(* Logix 5000 project; controller CIP vendor 1 type 14 code 106 rev 20.12; software revision 20.06; part 5 of 13 *)
(* tags used below, declared in another part *)
   Alarm_Ack : INT[8];
   Alarm_Present : INT[8];
   Alarm_Timer : TIMER[128];
   Bit : BOOL[128];
   IN_N7_100_199 : INT[100];
   Integer : DINT[150];
   OpCode_Pin : DINT[5];
   Recipe : RECIPE[41];
   RotaryONS : DINT;
   SCLD_Supply_Flow : REAL;
   SCLD_Supply_Pressure : REAL;
   SCLD_Wash_Chamber_Lvl : REAL;
   WashChamberDoorGasketCTRL : DINT;
(* MainProgram, continued *)

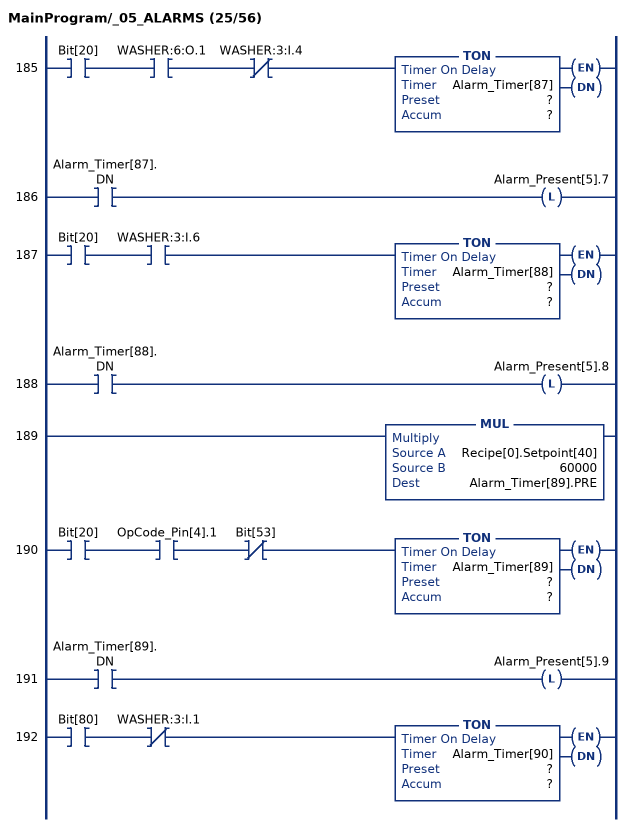
   [picture p67: MainProgram/_05_ALARMS rungs 185-192]
   185: XIC(Bit[20])XIC(WASHER:6:O.1)XIO(WASHER:3:I.4)TON(Alarm_Timer[87],?,?);
   186: XIC(Alarm_Timer[87].DN)OTL(Alarm_Present[5].7);
   187: XIC(Bit[20])XIC(WASHER:3:I.6)TON(Alarm_Timer[88],?,?);
   188: XIC(Alarm_Timer[88].DN)OTL(Alarm_Present[5].8);
   189: MUL(Recipe[0].Setpoint[40],60000,Alarm_Timer[89].PRE);
   190: XIC(Bit[20])XIC(OpCode_Pin[4].1)XIO(Bit[53])TON(Alarm_Timer[89],?,?);
   191: XIC(Alarm_Timer[89].DN)OTL(Alarm_Present[5].9);
   192: XIC(Bit[80])XIO(WASHER:3:I.1)TON(Alarm_Timer[90],?,?);
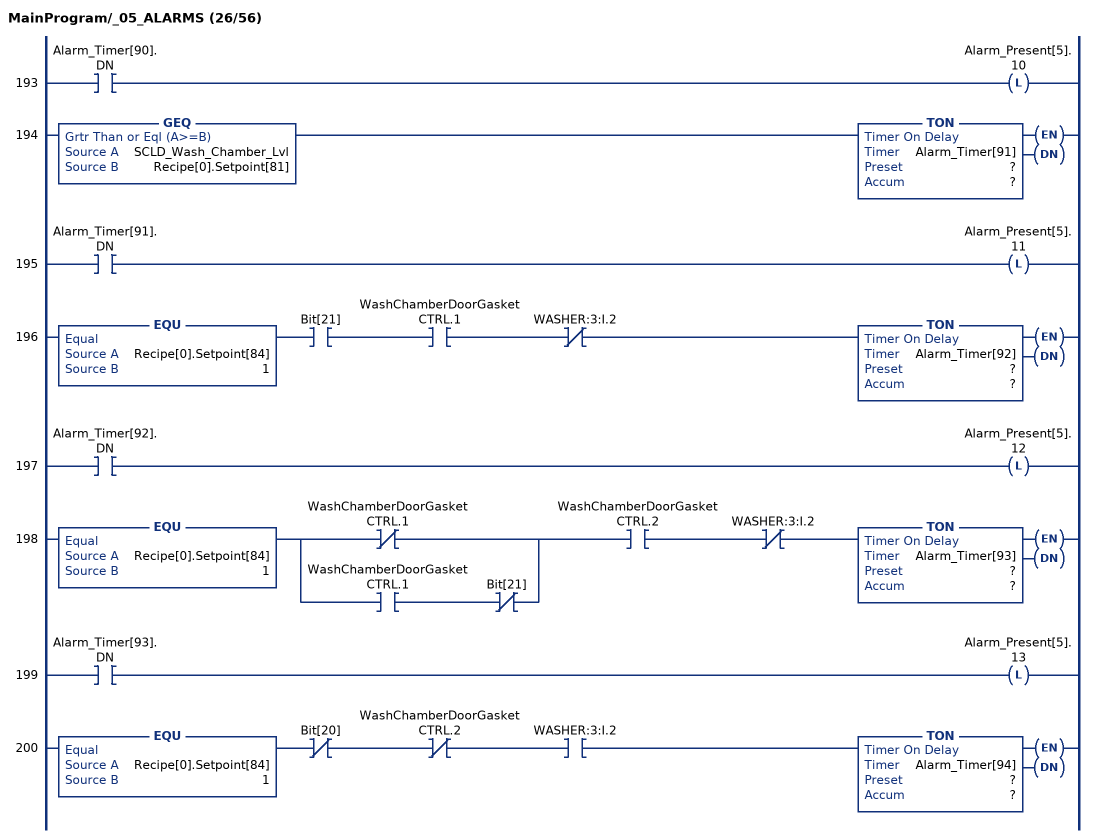
   193: XIC(Alarm_Timer[90].DN)OTL(Alarm_Present[5].10);
   194: GEQ(SCLD_Wash_Chamber_Lvl,Recipe[0].Setpoint[81])TON(Alarm_Timer[91],?,?);
   195: XIC(Alarm_Timer[91].DN)OTL(Alarm_Present[5].11);
   196: EQU(Recipe[0].Setpoint[84],1)XIC(Bit[21])XIC(WashChamberDoorGasketCTRL.1)XIO(WASHER:3:I.2)TON(Alarm_Timer[92],?,?);
   197: XIC(Alarm_Timer[92].DN)OTL(Alarm_Present[5].12);
   198: EQU(Recipe[0].Setpoint[84],1)[XIO(WashChamberDoorGasketCTRL.1) ,XIC(WashChamberDoorGasketCTRL.1) XIO(Bit[21]) ]XIC(WashChamberDoorGasketCTRL.2)XIO(WASHER:3:I.2)TON(Alarm_Timer[93],?,?);
   199: XIC(Alarm_Timer[93].DN)OTL(Alarm_Present[5].13);
   200: EQU(Recipe[0].Setpoint[84],1)XIO(Bit[20])XIO(WashChamberDoorGasketCTRL.2)XIC(WASHER:3:I.2)TON(Alarm_Timer[94],?,?);
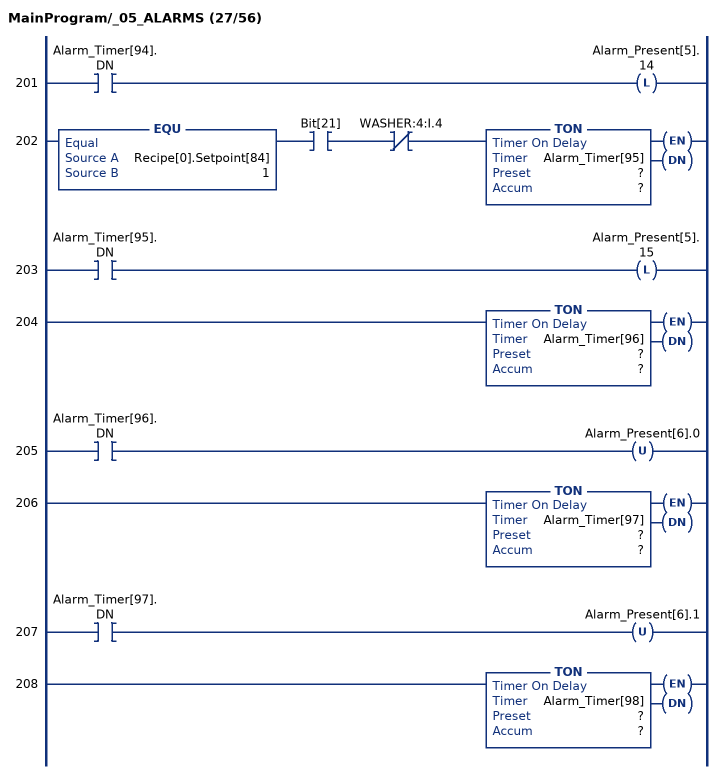
   201: XIC(Alarm_Timer[94].DN)OTL(Alarm_Present[5].14);
   202: EQU(Recipe[0].Setpoint[84],1)XIC(Bit[21])XIO(WASHER:4:I.4)TON(Alarm_Timer[95],?,?);
   203: XIC(Alarm_Timer[95].DN)OTL(Alarm_Present[5].15);
   204: TON(Alarm_Timer[96],?,?);
   205: XIC(Alarm_Timer[96].DN)OTU(Alarm_Present[6].0);
   206: TON(Alarm_Timer[97],?,?);
   207: XIC(Alarm_Timer[97].DN)OTU(Alarm_Present[6].1);
   208: TON(Alarm_Timer[98],?,?);
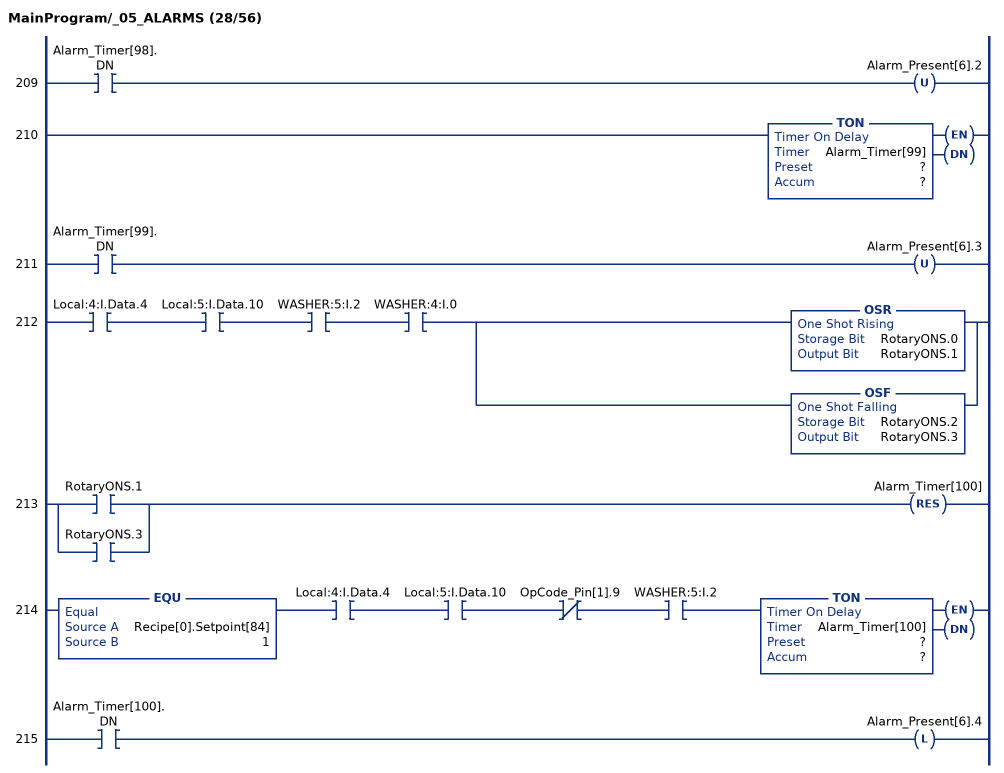
   209: XIC(Alarm_Timer[98].DN)OTU(Alarm_Present[6].2);
   210: TON(Alarm_Timer[99],?,?);
   211: XIC(Alarm_Timer[99].DN)OTU(Alarm_Present[6].3);
   212: XIC(Local:4:I.Data.4)XIC(Local:5:I.Data.10)XIC(WASHER:5:I.2)XIC(WASHER:4:I.0)[OSR(RotaryONS.0,RotaryONS.1) ,OSF(RotaryONS.2,RotaryONS.3) ];
   213: [XIC(RotaryONS.1) ,XIC(RotaryONS.3) ]RES(Alarm_Timer[100]);
   214: EQU(Recipe[0].Setpoint[84],1)XIC(Local:4:I.Data.4)XIC(Local:5:I.Data.10)XIO(OpCode_Pin[1].9)XIC(WASHER:5:I.2)TON(Alarm_Timer[100],?,?);
   215: XIC(Alarm_Timer[100].DN)OTL(Alarm_Present[6].4);
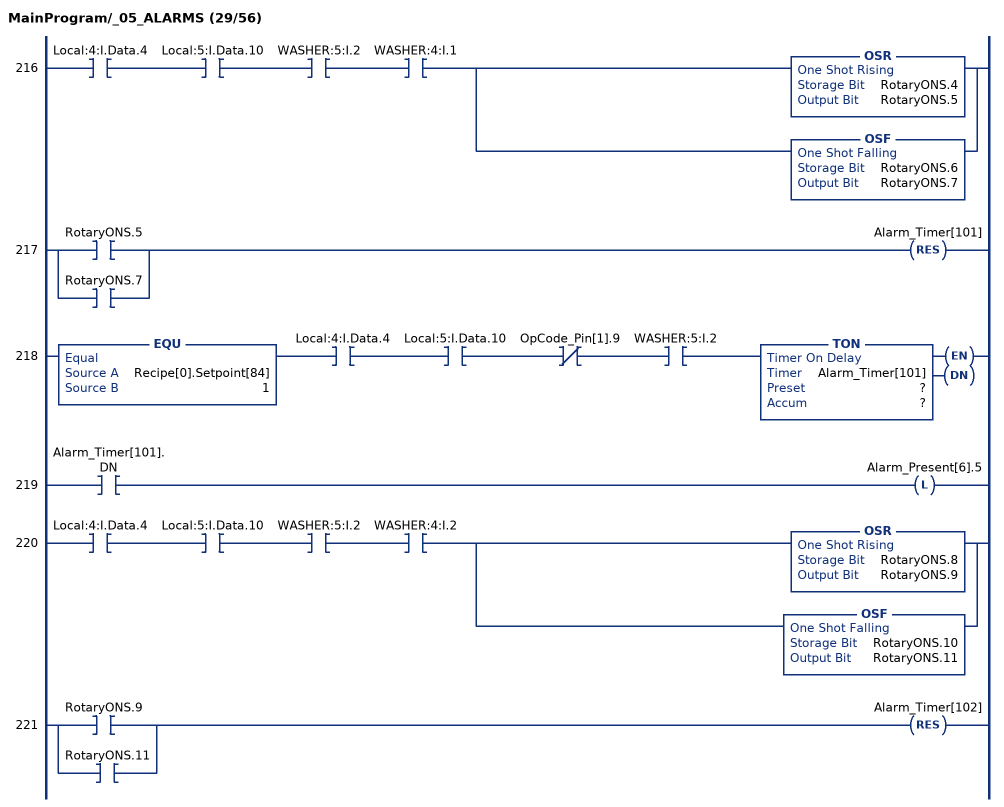
   216: XIC(Local:4:I.Data.4)XIC(Local:5:I.Data.10)XIC(WASHER:5:I.2)XIC(WASHER:4:I.1)[OSR(RotaryONS.4,RotaryONS.5) ,OSF(RotaryONS.6,RotaryONS.7) ];
   217: [XIC(RotaryONS.5) ,XIC(RotaryONS.7) ]RES(Alarm_Timer[101]);
   218: EQU(Recipe[0].Setpoint[84],1)XIC(Local:4:I.Data.4)XIC(Local:5:I.Data.10)XIO(OpCode_Pin[1].9)XIC(WASHER:5:I.2)TON(Alarm_Timer[101],?,?);
   219: XIC(Alarm_Timer[101].DN)OTL(Alarm_Present[6].5);
   220: XIC(Local:4:I.Data.4)XIC(Local:5:I.Data.10)XIC(WASHER:5:I.2)XIC(WASHER:4:I.2)[OSR(RotaryONS.8,RotaryONS.9) ,OSF(RotaryONS.10,RotaryONS.11) ];
   221: [XIC(RotaryONS.9) ,XIC(RotaryONS.11) ]RES(Alarm_Timer[102]);
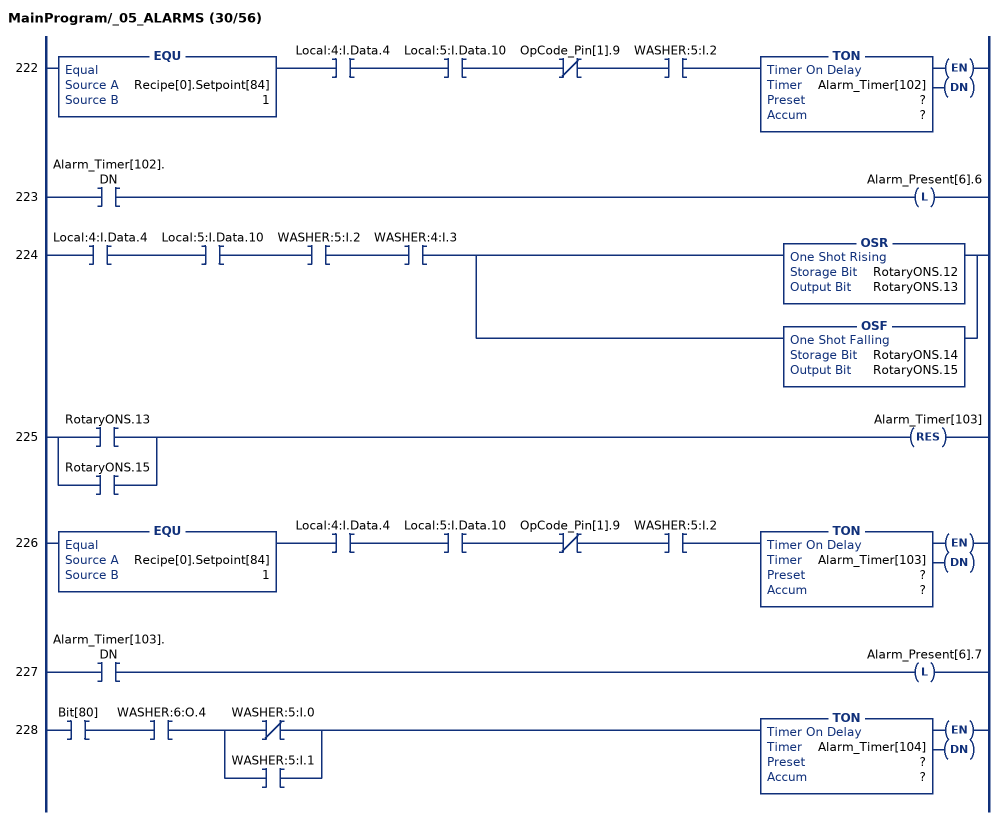
   222: EQU(Recipe[0].Setpoint[84],1)XIC(Local:4:I.Data.4)XIC(Local:5:I.Data.10)XIO(OpCode_Pin[1].9)XIC(WASHER:5:I.2)TON(Alarm_Timer[102],?,?);
   223: XIC(Alarm_Timer[102].DN)OTL(Alarm_Present[6].6);
   224: XIC(Local:4:I.Data.4)XIC(Local:5:I.Data.10)XIC(WASHER:5:I.2)XIC(WASHER:4:I.3)[OSR(RotaryONS.12,RotaryONS.13) ,OSF(RotaryONS.14,RotaryONS.15) ];
   225: [XIC(RotaryONS.13) ,XIC(RotaryONS.15) ]RES(Alarm_Timer[103]);
   226: EQU(Recipe[0].Setpoint[84],1)XIC(Local:4:I.Data.4)XIC(Local:5:I.Data.10)XIO(OpCode_Pin[1].9)XIC(WASHER:5:I.2)TON(Alarm_Timer[103],?,?);
   227: XIC(Alarm_Timer[103].DN)OTL(Alarm_Present[6].7);
   228: XIC(Bit[80])XIC(WASHER:6:O.4)[XIO(WASHER:5:I.0) ,XIC(WASHER:5:I.1) ]TON(Alarm_Timer[104],?,?);
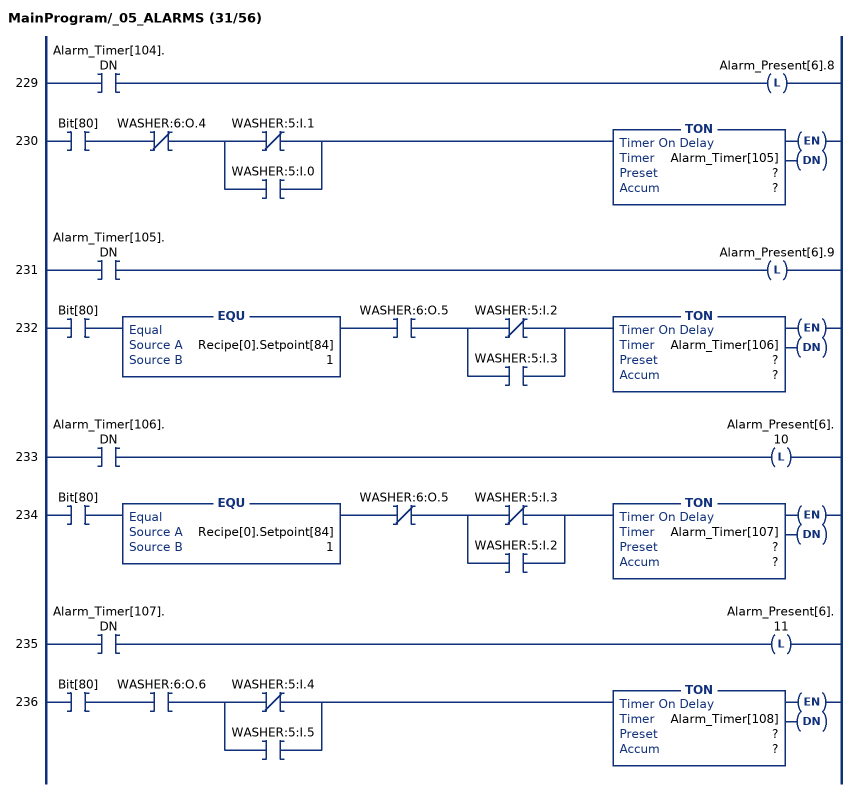
   229: XIC(Alarm_Timer[104].DN)OTL(Alarm_Present[6].8);
   230: XIC(Bit[80])XIO(WASHER:6:O.4)[XIO(WASHER:5:I.1) ,XIC(WASHER:5:I.0) ]TON(Alarm_Timer[105],?,?);
   231: XIC(Alarm_Timer[105].DN)OTL(Alarm_Present[6].9);
   232: XIC(Bit[80])EQU(Recipe[0].Setpoint[84],1)XIC(WASHER:6:O.5)[XIO(WASHER:5:I.2) ,XIC(WASHER:5:I.3) ]TON(Alarm_Timer[106],?,?);
   233: XIC(Alarm_Timer[106].DN)OTL(Alarm_Present[6].10);
   234: XIC(Bit[80])EQU(Recipe[0].Setpoint[84],1)XIO(WASHER:6:O.5)[XIO(WASHER:5:I.3) ,XIC(WASHER:5:I.2) ]TON(Alarm_Timer[107],?,?);
   235: XIC(Alarm_Timer[107].DN)OTL(Alarm_Present[6].11);
   236: XIC(Bit[80])XIC(WASHER:6:O.6)[XIO(WASHER:5:I.4) ,XIC(WASHER:5:I.5) ]TON(Alarm_Timer[108],?,?);
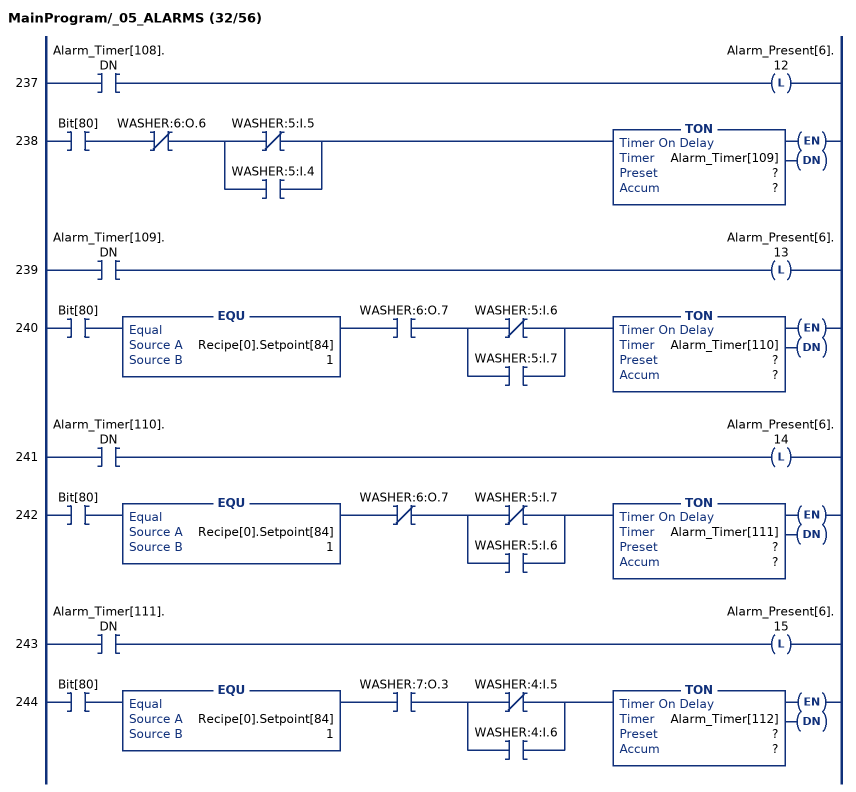
   237: XIC(Alarm_Timer[108].DN)OTL(Alarm_Present[6].12);
   238: XIC(Bit[80])XIO(WASHER:6:O.6)[XIO(WASHER:5:I.5) ,XIC(WASHER:5:I.4) ]TON(Alarm_Timer[109],?,?);
   239: XIC(Alarm_Timer[109].DN)OTL(Alarm_Present[6].13);
   240: XIC(Bit[80])EQU(Recipe[0].Setpoint[84],1)XIC(WASHER:6:O.7)[XIO(WASHER:5:I.6) ,XIC(WASHER:5:I.7) ]TON(Alarm_Timer[110],?,?);
   241: XIC(Alarm_Timer[110].DN)OTL(Alarm_Present[6].14);
   242: XIC(Bit[80])EQU(Recipe[0].Setpoint[84],1)XIO(WASHER:6:O.7)[XIO(WASHER:5:I.7) ,XIC(WASHER:5:I.6) ]TON(Alarm_Timer[111],?,?);
   243: XIC(Alarm_Timer[111].DN)OTL(Alarm_Present[6].15);
   244: XIC(Bit[80])EQU(Recipe[0].Setpoint[84],1)XIC(WASHER:7:O.3)[XIO(WASHER:4:I.5) ,XIC(WASHER:4:I.6) ]TON(Alarm_Timer[112],?,?);
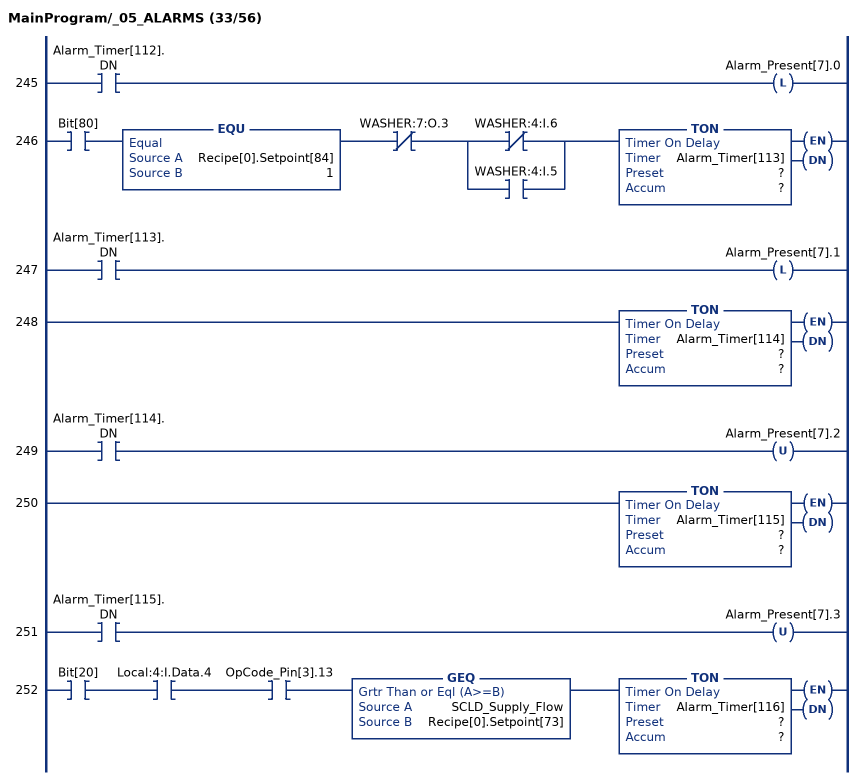
   245: XIC(Alarm_Timer[112].DN)OTL(Alarm_Present[7].0);
   246: XIC(Bit[80])EQU(Recipe[0].Setpoint[84],1)XIO(WASHER:7:O.3)[XIO(WASHER:4:I.6) ,XIC(WASHER:4:I.5) ]TON(Alarm_Timer[113],?,?);
   247: XIC(Alarm_Timer[113].DN)OTL(Alarm_Present[7].1);
   248: TON(Alarm_Timer[114],?,?);
   249: XIC(Alarm_Timer[114].DN)OTU(Alarm_Present[7].2);
   250: TON(Alarm_Timer[115],?,?);
   251: XIC(Alarm_Timer[115].DN)OTU(Alarm_Present[7].3);
   252: XIC(Bit[20])XIC(Local:4:I.Data.4)XIC(OpCode_Pin[3].13)GEQ(SCLD_Supply_Flow,Recipe[0].Setpoint[73])TON(Alarm_Timer[116],?,?);
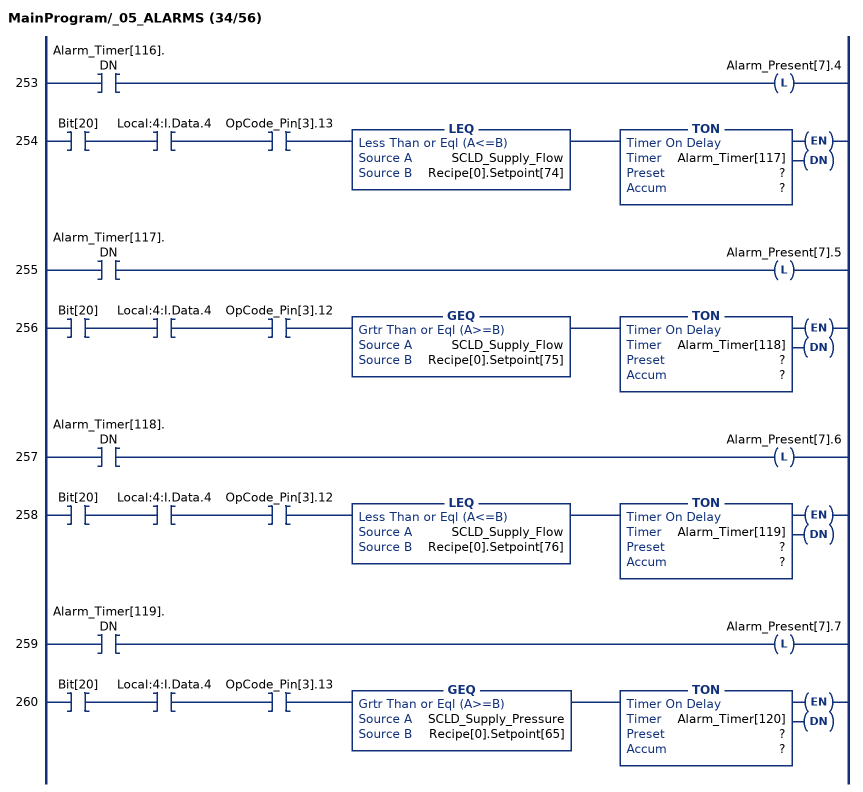
   253: XIC(Alarm_Timer[116].DN)OTL(Alarm_Present[7].4);
   254: XIC(Bit[20])XIC(Local:4:I.Data.4)XIC(OpCode_Pin[3].13)LEQ(SCLD_Supply_Flow,Recipe[0].Setpoint[74])TON(Alarm_Timer[117],?,?);
   255: XIC(Alarm_Timer[117].DN)OTL(Alarm_Present[7].5);
   256: XIC(Bit[20])XIC(Local:4:I.Data.4)XIC(OpCode_Pin[3].12)GEQ(SCLD_Supply_Flow,Recipe[0].Setpoint[75])TON(Alarm_Timer[118],?,?);
   257: XIC(Alarm_Timer[118].DN)OTL(Alarm_Present[7].6);
   258: XIC(Bit[20])XIC(Local:4:I.Data.4)XIC(OpCode_Pin[3].12)LEQ(SCLD_Supply_Flow,Recipe[0].Setpoint[76])TON(Alarm_Timer[119],?,?);
   259: XIC(Alarm_Timer[119].DN)OTL(Alarm_Present[7].7);
   260: XIC(Bit[20])XIC(Local:4:I.Data.4)XIC(OpCode_Pin[3].13)GEQ(SCLD_Supply_Pressure,Recipe[0].Setpoint[65])TON(Alarm_Timer[120],?,?);
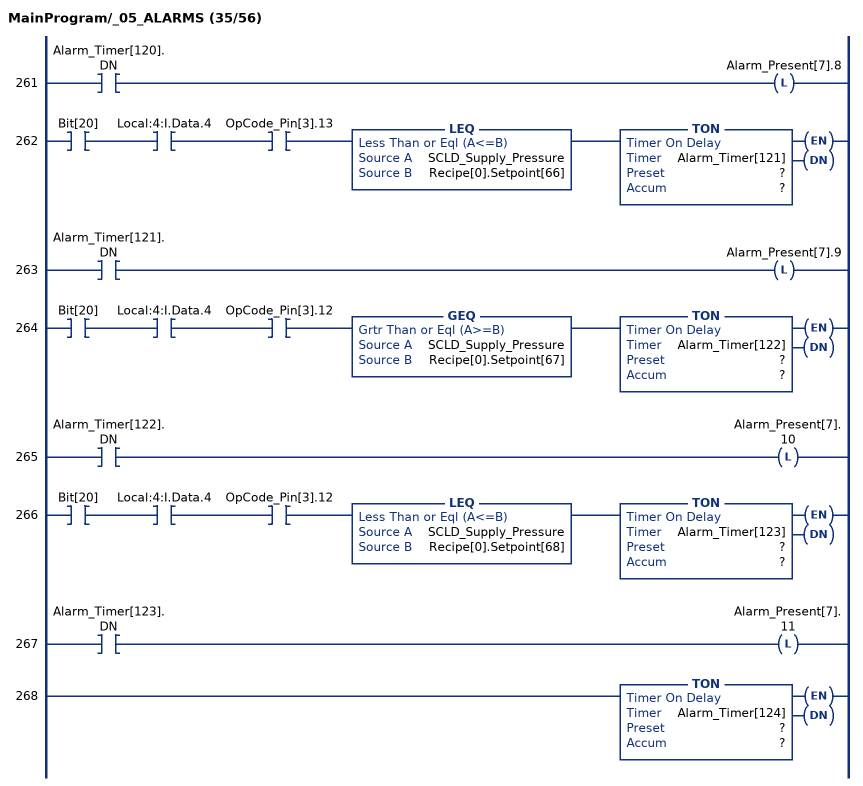
   261: XIC(Alarm_Timer[120].DN)OTL(Alarm_Present[7].8);
   262: XIC(Bit[20])XIC(Local:4:I.Data.4)XIC(OpCode_Pin[3].13)LEQ(SCLD_Supply_Pressure,Recipe[0].Setpoint[66])TON(Alarm_Timer[121],?,?);
   263: XIC(Alarm_Timer[121].DN)OTL(Alarm_Present[7].9);
   264: XIC(Bit[20])XIC(Local:4:I.Data.4)XIC(OpCode_Pin[3].12)GEQ(SCLD_Supply_Pressure,Recipe[0].Setpoint[67])TON(Alarm_Timer[122],?,?);
   265: XIC(Alarm_Timer[122].DN)OTL(Alarm_Present[7].10);
   266: XIC(Bit[20])XIC(Local:4:I.Data.4)XIC(OpCode_Pin[3].12)LEQ(SCLD_Supply_Pressure,Recipe[0].Setpoint[68])TON(Alarm_Timer[123],?,?);
   267: XIC(Alarm_Timer[123].DN)OTL(Alarm_Present[7].11);
   268: TON(Alarm_Timer[124],?,?);
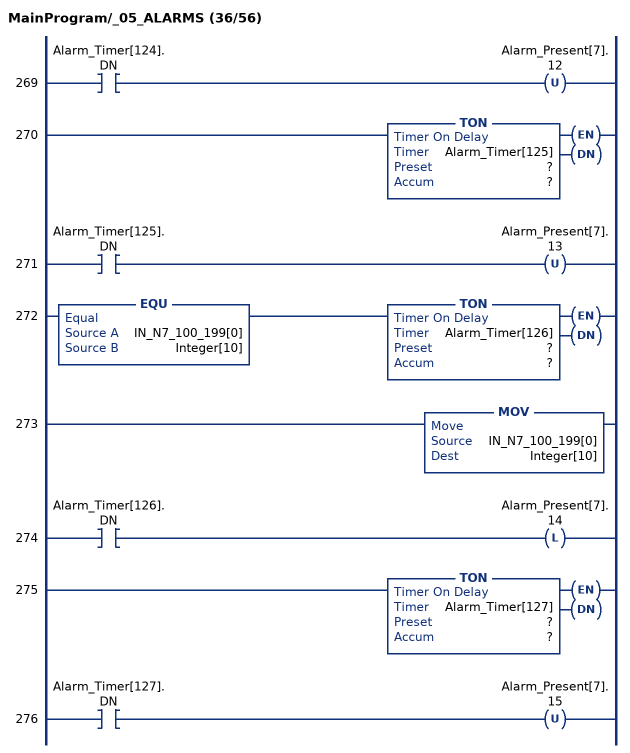
   269: XIC(Alarm_Timer[124].DN)OTU(Alarm_Present[7].12);
   270: TON(Alarm_Timer[125],?,?);
   271: XIC(Alarm_Timer[125].DN)OTU(Alarm_Present[7].13);
   272: EQU(IN_N7_100_199[0],Integer[10])TON(Alarm_Timer[126],?,?);
   273: MOV(IN_N7_100_199[0],Integer[10]);
   274: XIC(Alarm_Timer[126].DN)OTL(Alarm_Present[7].14);
   275: TON(Alarm_Timer[127],?,?);
   276: XIC(Alarm_Timer[127].DN)OTU(Alarm_Present[7].15);
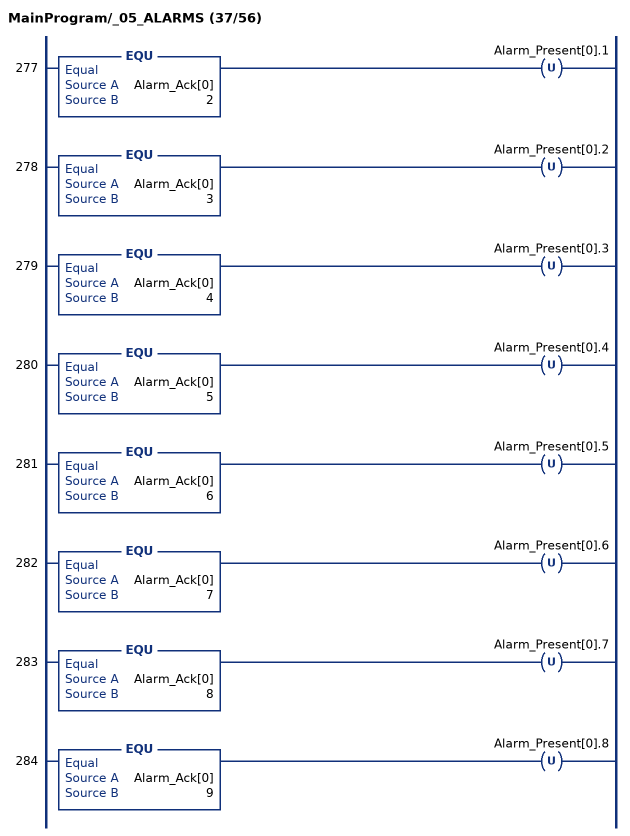
   277: EQU(Alarm_Ack[0],2)OTU(Alarm_Present[0].1);
   278: EQU(Alarm_Ack[0],3)OTU(Alarm_Present[0].2);
   279: EQU(Alarm_Ack[0],4)OTU(Alarm_Present[0].3);
   280: EQU(Alarm_Ack[0],5)OTU(Alarm_Present[0].4);
   281: EQU(Alarm_Ack[0],6)OTU(Alarm_Present[0].5);
   282: EQU(Alarm_Ack[0],7)OTU(Alarm_Present[0].6);
   283: EQU(Alarm_Ack[0],8)OTU(Alarm_Present[0].7);
   284: EQU(Alarm_Ack[0],9)OTU(Alarm_Present[0].8);
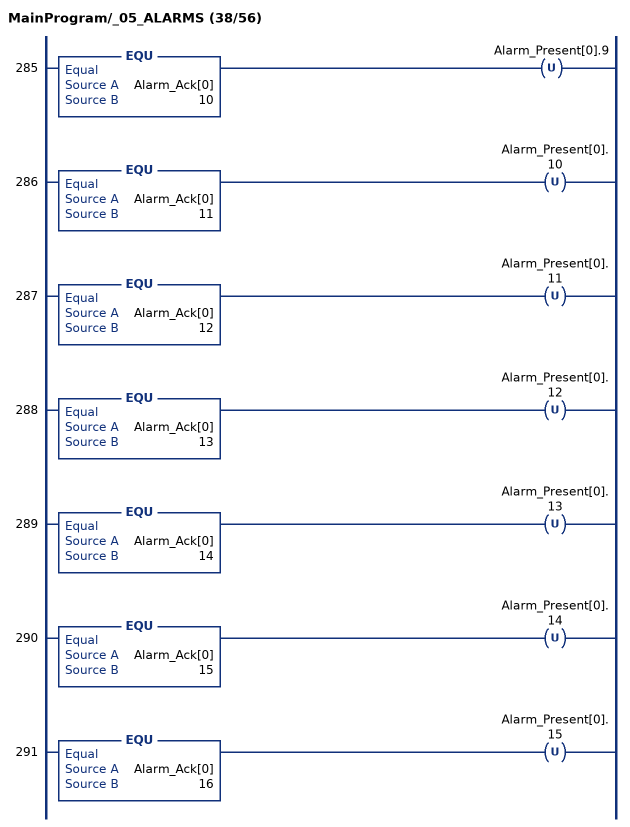
   285: EQU(Alarm_Ack[0],10)OTU(Alarm_Present[0].9);
   286: EQU(Alarm_Ack[0],11)OTU(Alarm_Present[0].10);
   287: EQU(Alarm_Ack[0],12)OTU(Alarm_Present[0].11);
   288: EQU(Alarm_Ack[0],13)OTU(Alarm_Present[0].12);
   289: EQU(Alarm_Ack[0],14)OTU(Alarm_Present[0].13);
   290: EQU(Alarm_Ack[0],15)OTU(Alarm_Present[0].14);
   291: EQU(Alarm_Ack[0],16)OTU(Alarm_Present[0].15);
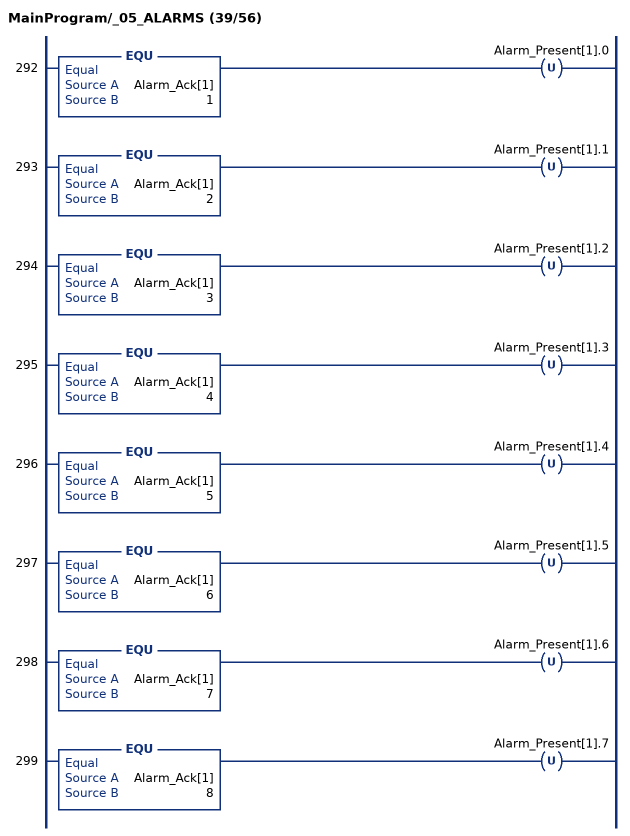
   292: EQU(Alarm_Ack[1],1)OTU(Alarm_Present[1].0);
   293: EQU(Alarm_Ack[1],2)OTU(Alarm_Present[1].1);
   294: EQU(Alarm_Ack[1],3)OTU(Alarm_Present[1].2);
   295: EQU(Alarm_Ack[1],4)OTU(Alarm_Present[1].3);
   296: EQU(Alarm_Ack[1],5)OTU(Alarm_Present[1].4);
   297: EQU(Alarm_Ack[1],6)OTU(Alarm_Present[1].5);
   298: EQU(Alarm_Ack[1],7)OTU(Alarm_Present[1].6);
   299: EQU(Alarm_Ack[1],8)OTU(Alarm_Present[1].7);
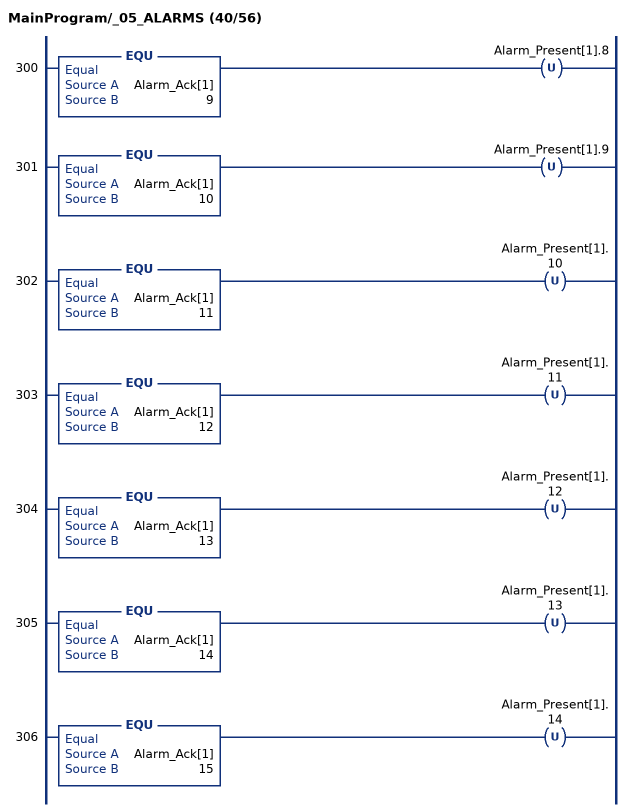
   300: EQU(Alarm_Ack[1],9)OTU(Alarm_Present[1].8);
   301: EQU(Alarm_Ack[1],10)OTU(Alarm_Present[1].9);
   302: EQU(Alarm_Ack[1],11)OTU(Alarm_Present[1].10);
   303: EQU(Alarm_Ack[1],12)OTU(Alarm_Present[1].11);
   304: EQU(Alarm_Ack[1],13)OTU(Alarm_Present[1].12);
   305: EQU(Alarm_Ack[1],14)OTU(Alarm_Present[1].13);
   306: EQU(Alarm_Ack[1],15)OTU(Alarm_Present[1].14);
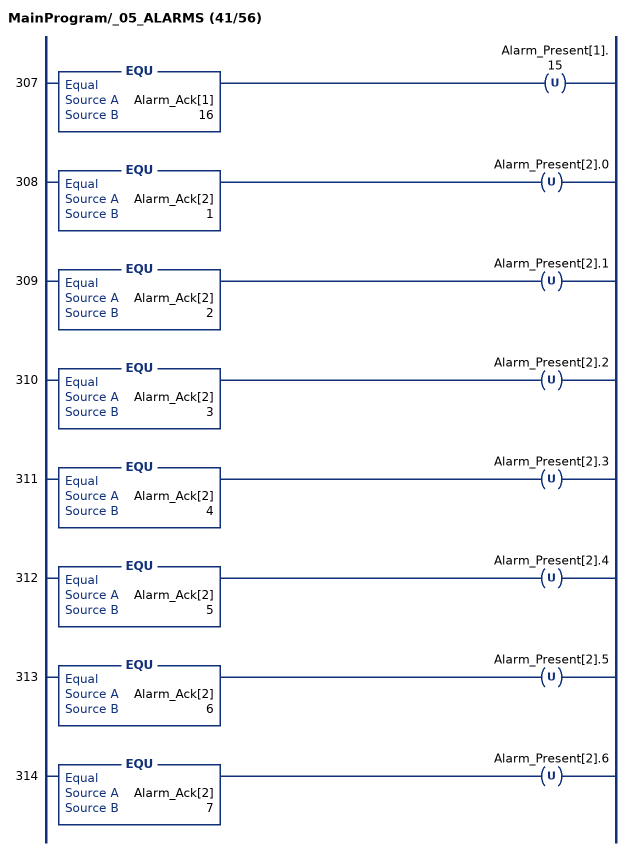
   307: EQU(Alarm_Ack[1],16)OTU(Alarm_Present[1].15);
   308: EQU(Alarm_Ack[2],1)OTU(Alarm_Present[2].0);
   309: EQU(Alarm_Ack[2],2)OTU(Alarm_Present[2].1);
   310: EQU(Alarm_Ack[2],3)OTU(Alarm_Present[2].2);
   311: EQU(Alarm_Ack[2],4)OTU(Alarm_Present[2].3);
   312: EQU(Alarm_Ack[2],5)OTU(Alarm_Present[2].4);
   313: EQU(Alarm_Ack[2],6)OTU(Alarm_Present[2].5);
   314: EQU(Alarm_Ack[2],7)OTU(Alarm_Present[2].6);
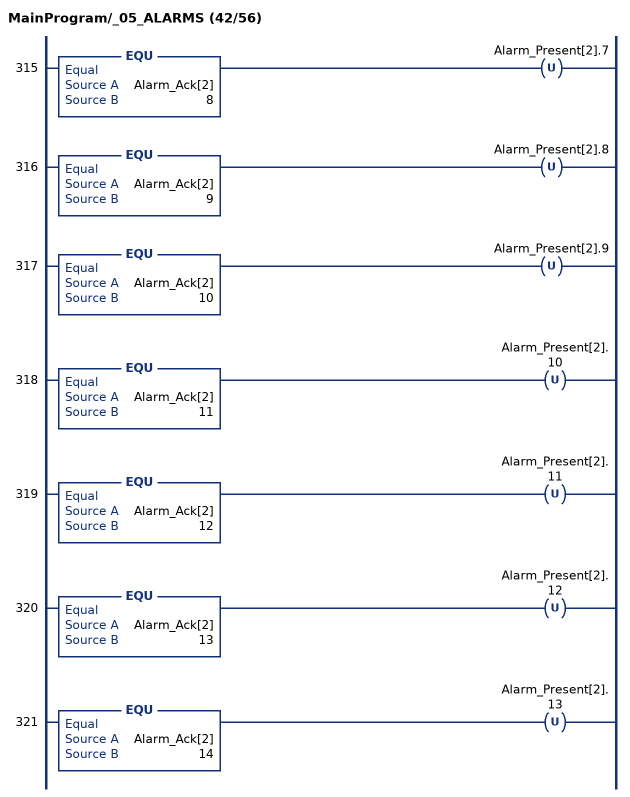
   315: EQU(Alarm_Ack[2],8)OTU(Alarm_Present[2].7);
   316: EQU(Alarm_Ack[2],9)OTU(Alarm_Present[2].8);
   317: EQU(Alarm_Ack[2],10)OTU(Alarm_Present[2].9);
   318: EQU(Alarm_Ack[2],11)OTU(Alarm_Present[2].10);
   319: EQU(Alarm_Ack[2],12)OTU(Alarm_Present[2].11);
   320: EQU(Alarm_Ack[2],13)OTU(Alarm_Present[2].12);
   321: EQU(Alarm_Ack[2],14)OTU(Alarm_Present[2].13);
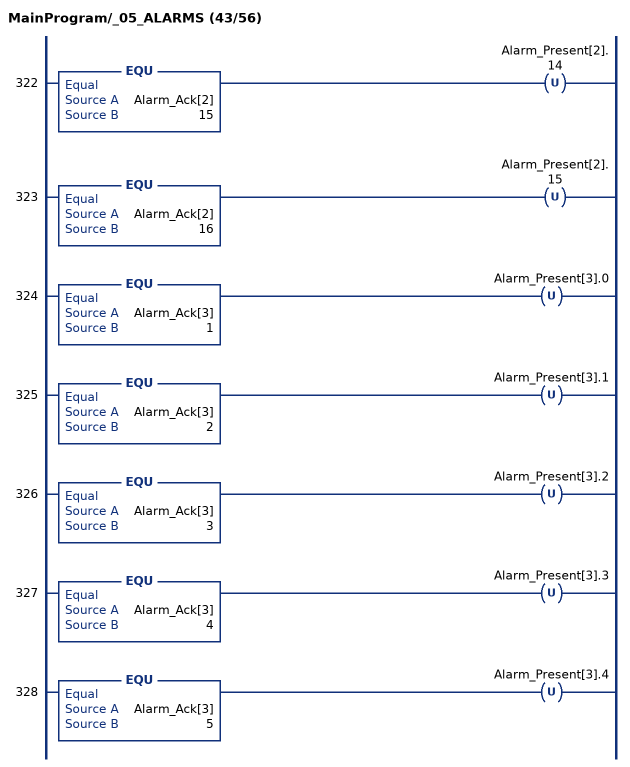
   322: EQU(Alarm_Ack[2],15)OTU(Alarm_Present[2].14);
   323: EQU(Alarm_Ack[2],16)OTU(Alarm_Present[2].15);
   324: EQU(Alarm_Ack[3],1)OTU(Alarm_Present[3].0);
   325: EQU(Alarm_Ack[3],2)OTU(Alarm_Present[3].1);
   326: EQU(Alarm_Ack[3],3)OTU(Alarm_Present[3].2);
   327: EQU(Alarm_Ack[3],4)OTU(Alarm_Present[3].3);
   328: EQU(Alarm_Ack[3],5)OTU(Alarm_Present[3].4);
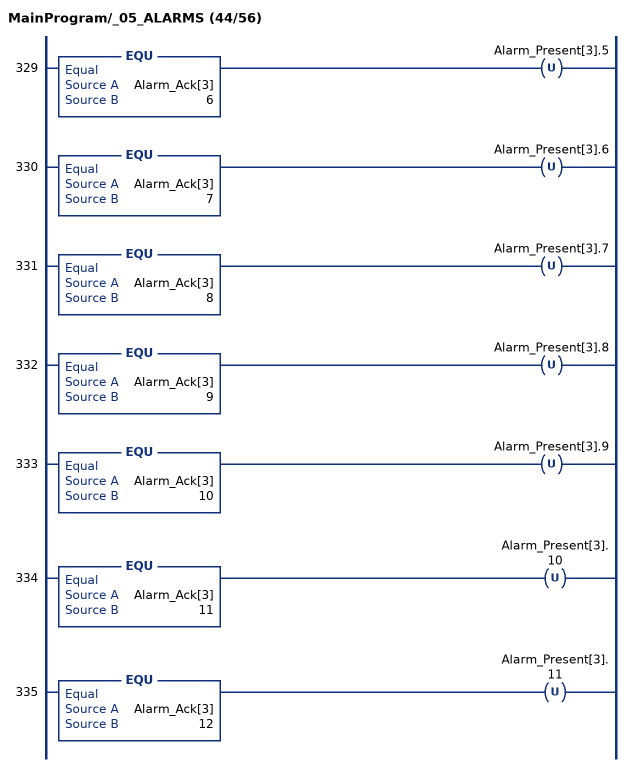
   329: EQU(Alarm_Ack[3],6)OTU(Alarm_Present[3].5);
   330: EQU(Alarm_Ack[3],7)OTU(Alarm_Present[3].6);
   331: EQU(Alarm_Ack[3],8)OTU(Alarm_Present[3].7);
   332: EQU(Alarm_Ack[3],9)OTU(Alarm_Present[3].8);
   333: EQU(Alarm_Ack[3],10)OTU(Alarm_Present[3].9);
   334: EQU(Alarm_Ack[3],11)OTU(Alarm_Present[3].10);
   335: EQU(Alarm_Ack[3],12)OTU(Alarm_Present[3].11);
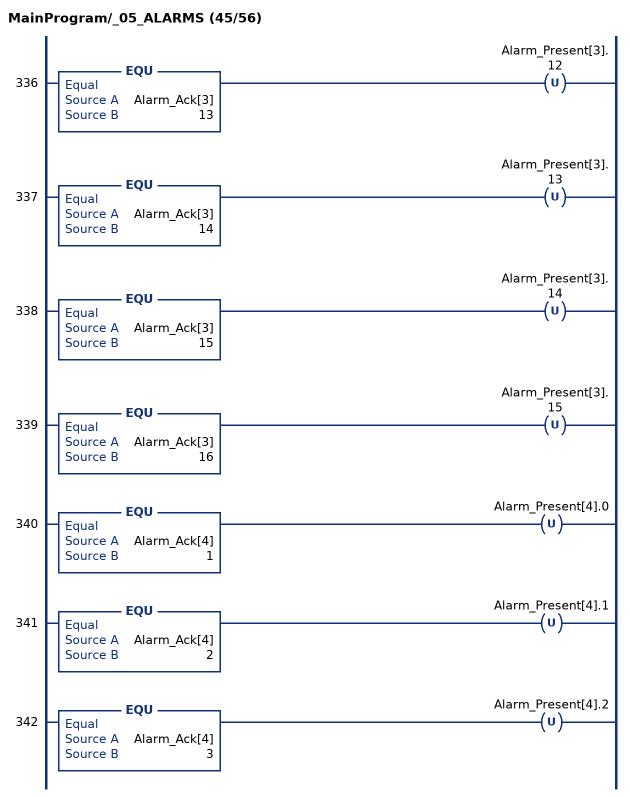
   336: EQU(Alarm_Ack[3],13)OTU(Alarm_Present[3].12);
   337: EQU(Alarm_Ack[3],14)OTU(Alarm_Present[3].13);
   338: EQU(Alarm_Ack[3],15)OTU(Alarm_Present[3].14);
   339: EQU(Alarm_Ack[3],16)OTU(Alarm_Present[3].15);
   340: EQU(Alarm_Ack[4],1)OTU(Alarm_Present[4].0);
   341: EQU(Alarm_Ack[4],2)OTU(Alarm_Present[4].1);
   342: EQU(Alarm_Ack[4],3)OTU(Alarm_Present[4].2);
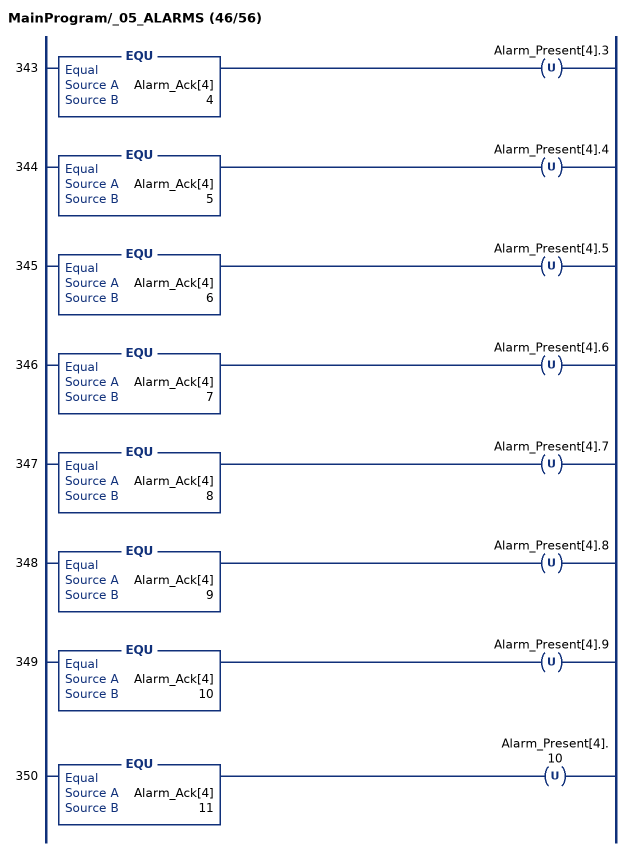
   343: EQU(Alarm_Ack[4],4)OTU(Alarm_Present[4].3);
   344: EQU(Alarm_Ack[4],5)OTU(Alarm_Present[4].4);
   345: EQU(Alarm_Ack[4],6)OTU(Alarm_Present[4].5);
   346: EQU(Alarm_Ack[4],7)OTU(Alarm_Present[4].6);
   347: EQU(Alarm_Ack[4],8)OTU(Alarm_Present[4].7);
   348: EQU(Alarm_Ack[4],9)OTU(Alarm_Present[4].8);
   349: EQU(Alarm_Ack[4],10)OTU(Alarm_Present[4].9);
   350: EQU(Alarm_Ack[4],11)OTU(Alarm_Present[4].10);
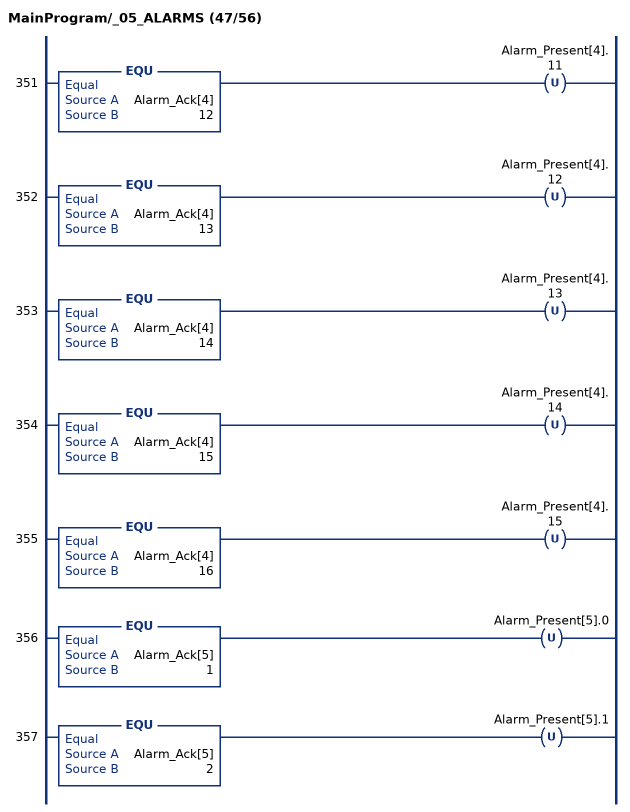
   351: EQU(Alarm_Ack[4],12)OTU(Alarm_Present[4].11);
   352: EQU(Alarm_Ack[4],13)OTU(Alarm_Present[4].12);
   353: EQU(Alarm_Ack[4],14)OTU(Alarm_Present[4].13);
   354: EQU(Alarm_Ack[4],15)OTU(Alarm_Present[4].14);
   355: EQU(Alarm_Ack[4],16)OTU(Alarm_Present[4].15);
   356: EQU(Alarm_Ack[5],1)OTU(Alarm_Present[5].0);
   357: EQU(Alarm_Ack[5],2)OTU(Alarm_Present[5].1);
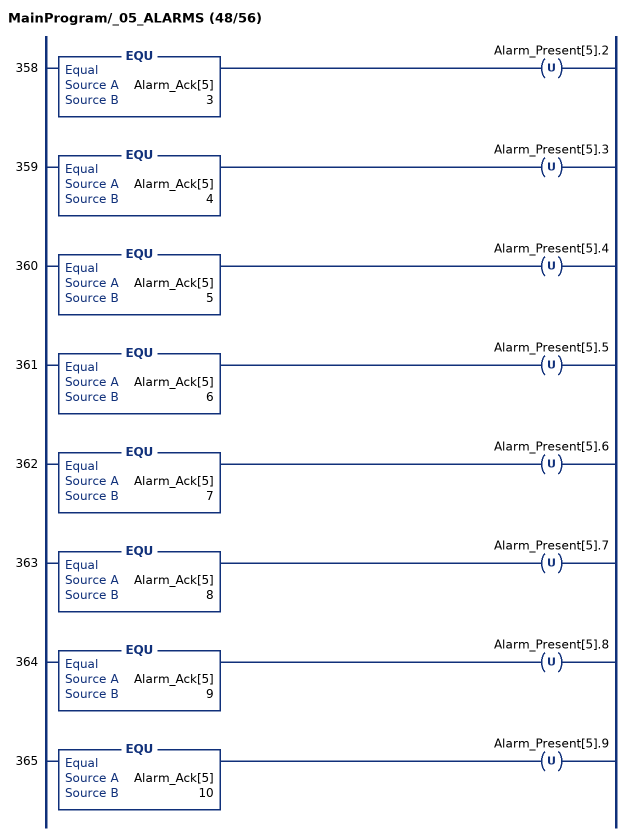
   358: EQU(Alarm_Ack[5],3)OTU(Alarm_Present[5].2);
   359: EQU(Alarm_Ack[5],4)OTU(Alarm_Present[5].3);
   360: EQU(Alarm_Ack[5],5)OTU(Alarm_Present[5].4);
   361: EQU(Alarm_Ack[5],6)OTU(Alarm_Present[5].5);
   362: EQU(Alarm_Ack[5],7)OTU(Alarm_Present[5].6);
   363: EQU(Alarm_Ack[5],8)OTU(Alarm_Present[5].7);
   364: EQU(Alarm_Ack[5],9)OTU(Alarm_Present[5].8);
   365: EQU(Alarm_Ack[5],10)OTU(Alarm_Present[5].9);
